(* IEC 61131-3 sources: sis-interlock-demo/tools/tests/fixtures/sample/src/POUs/Devices/FB_Motor, 5 files *)

(* ---- FB_Motor.decl.st ---- *)
(*
    Назначение: двигатель с контактором — пуск, стоп, контроль обратной связи
    Автор: kr0nsch
    Версия: 1.0.0
    Документ: docs/ARCHITECTURE.md
*)
FUNCTION_BLOCK FB_Motor EXTENDS FB_DeviceBase
VAR_INPUT
    stCmd : ST_MotorCmd;            // команды HMI
    xFeedback : BOOL;               // обратная связь контактора
    itfInterlock : I_Resettable;    // связанная блокировка (необязательно)
END_VAR
VAR_OUTPUT
    xRun : BOOL;                    // команда на контактор
    stSts : ST_MotorSts;            // состояние для HMI
END_VAR
VAR
    fbStartTimer : TON;             // контроль обратной связи при пуске
    fbAckEdge : R_TRIG;             // фронт квитирования
    rSpeedSp_rpm : REAL;            // принятая уставка
    pSts : POINTER TO ST_MotorSts;
    refCmd : REFERENCE TO ST_MotorCmd;
    iStep : INT := GVL_Const.STEP_IDLE;
    wsState : WSTRING(80) := "Остановлен";
END_VAR

(* ---- FB_Motor.impl.st ---- *)
refCmd REF= stCmd;
pSts := ADR(stSts);
fbAckEdge(CLK := refCmd.xAck);
IF fbAckEdge.Q THEN
    Reset(xForce := FALSE);
END_IF

CASE eModeInt OF
    E_DeviceMode.Auto, E_DeviceMode.Manual:
        IF refCmd.xStart AND xEnable AND NOT xFault THEN
            xRun := TRUE;
            iStep := GVL_Const.STEP_RUN;
        END_IF
    E_DeviceMode.OutOfService:
        xRun := FALSE;
ELSE
    xRun := FALSE;
END_CASE
xRun R= refCmd.xStop OR xFault;

CASE iStep OF
    GVL_Const.STEP_IDLE:
        wsState := "Остановлен";
    GVL_Const.STEP_RUN:
        wsState := "В работе";
END_CASE

(* Нет обратной связи за MOTOR_START_TIMEOUT — отказ *)
fbStartTimer(IN := xRun AND NOT xFeedback, PT := GVL_Const.MOTOR_START_TIMEOUT);
xFault S= fbStartTimer.Q;
IF xFault THEN
    eNamur := E_NamurStatus.Failure;
    wsState := "Авария: нет обратной связи";
END_IF

pSts^.xRunning := xRun AND xFeedback;
pSts^.xFault := xFault;
stSts.eMode := eModeInt;
stSts.eNamur := eNamur;
stSts.rSpeed_rpm := F_Clamp(
    rValue := rSpeedSp_rpm,
    rMin := GVL_Const.MOTOR_SPEED_MIN_RPM,
    rMax := GVL_Const.MOTOR_SPEED_MAX_RPM);
stSts.wsText := wsState;

(* ---- Reset.method.decl.st ---- *)
METHOD PUBLIC Reset : BOOL
VAR_INPUT
    xForce : BOOL;
END_VAR

(* ---- Reset.method.impl.st ---- *)
Reset := SUPER^.Reset(xForce := xForce);
IF itfInterlock <> 0 THEN
    itfInterlock.Reset(xForce := xForce);
END_IF
fbStartTimer(IN := FALSE);
iStep := GVL_Const.STEP_IDLE;

(* ---- Start.method.decl.st ---- *)
METHOD PUBLIC Start
VAR_INPUT
    rSpeed_rpm : REAL;
END_VAR
